SUBAPPLICATION AUDI_GT_0 (* Prüft ob UDINT-Adapter Wert > 0 ist (AX-Adapter Ausgang) *)
  (* Standard: 61499-2 *)
  (* Version 1.0, 2026-10-15, franz, Meisterschulen am Ostbahnhof *)
  PACKAGE MyLib::sys;
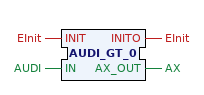
  EVENT_INPUT
    INIT : EInit; (* Initialization Request *)
  END_EVENT
  EVENT_OUTPUT
    INITO : EInit; (* Initialization Confirm *)
  END_EVENT
  SOCKETS
    IN : adapter::types::unidirectional::AUDI;
  END_SOCKETS
  PLUGS
    AX_OUT : adapter::types::unidirectional::AX;
  END_PLUGS
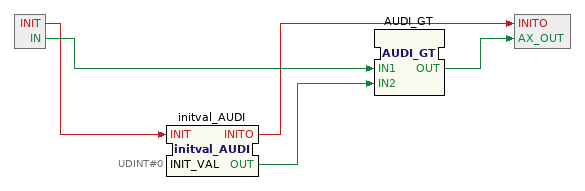
  FBS
    AUDI_GT : adapter::iec61131::comparison::AUDI_GT;
    initval_AUDI : adapter::types::unidirectional::AUDI::initval::initval_AUDI(INIT_VAL := UDINT#0);
  END_FBS
  EVENT_CONNECTIONS
    INIT TO initval_AUDI.INIT;
    initval_AUDI.INITO TO INITO;
  END_CONNECTIONS
  ADAPTER_CONNECTIONS
    IN TO AUDI_GT.IN1;
    AUDI_GT.OUT TO AX_OUT;
    initval_AUDI.OUT TO AUDI_GT.IN2;
  END_CONNECTIONS
END_SUBAPPLICATION
